# EPICS substitutions: b-55B2VNC/src/main/epics/PCF0CoreApp/Db/nisyncDevice6683H-terminal.substitutions
#TERMINAL 0-18
file "./nisync_Terminal.template" {
pattern {BOARDTYPE,	BOARDTYPEIDX,	CBS1,	CBS2,	TERMINAL_NAME}
		{"B",		"1",			"D1",	"I2",	"TR0" }
		{"B",		"1",			"D1",	"I2",	"TR1" }
		{"B",		"1",			"D1",	"I2",	"TR2" }
		{"B",		"1",			"D1",	"I2",	"TR11"}
		{"B",		"1",			"D1",	"I2",	"TR12"}
		{"B",		"1",			"D1",	"I2",	"TR13"}
		{"B",		"1",			"D1",	"I2",	"TR14"}
		{"B",		"1",			"D1",	"I2",	"TR15"}
		{"B",		"1",			"D1",	"I2",	"TR16"}
		{"B",		"1",			"D1",	"I2",	"TR17"}
		{"B",		"1",			"D1",	"I2",	"TR18"}

}
